{attribute 'qualified_only'}
{attribute 'to_string'}
TYPE E_Anybus_ClientType :
(
	eNone	:= 0,	// not selected
	ePipe	:= 1,	// no spray ball
	eTank	:= 2	// always with a spray ball, decided 01.11.2026
);
END_TYPE

(* stored: Version 1.1.0.1, ProductVersion 3.1.4026.20
   DUT E_Anybus_ClientType: Id {e066ad1d-5a6d-4bc4-9863-2ec5626c1e3f} *)
